FUNCTION_BLOCK GATE_CYCLE
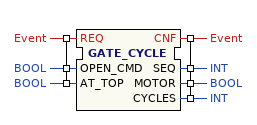
  EVENT_INPUT
    REQ WITH OPEN_CMD, AT_TOP;
  END_EVENT
  EVENT_OUTPUT
    CNF WITH SEQ, MOTOR, CYCLES;
  END_EVENT
  VAR_INPUT
    OPEN_CMD : BOOL;
    AT_TOP : BOOL;
  END_VAR
  VAR_OUTPUT
    SEQ : INT;
    MOTOR : BOOL;
    CYCLES : INT;
  END_VAR
  VAR
    SEQ_STATE : INT;
    SEQ_START_TIME : TIME;
  END_VAR
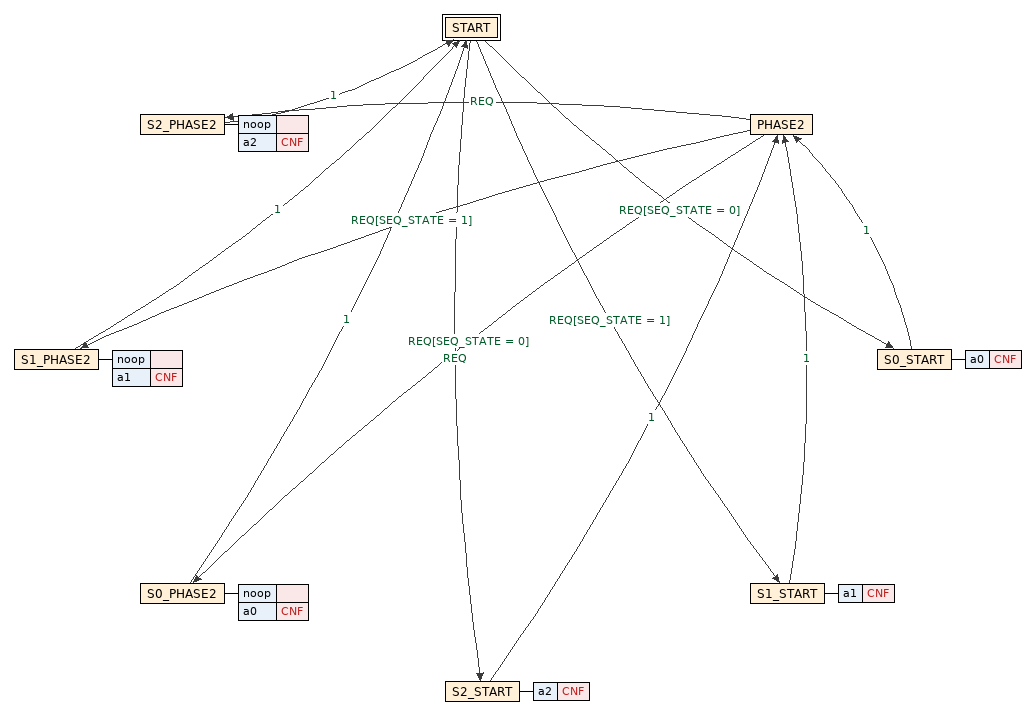
  EC_STATES
    START;
    PHASE2;
    S0_START : a0 -> CNF;
    S1_START : a1 -> CNF;
    S2_START : a2 -> CNF;
    S0_PHASE2 : noop, a0 -> CNF;
    S1_PHASE2 : noop, a1 -> CNF;
    S2_PHASE2 : noop, a2 -> CNF;
  END_STATES
  EC_TRANSITIONS
    START TO S0_START := REQ[SEQ_STATE = 0];
    START TO S1_START := REQ[SEQ_STATE = 1];
    START TO S2_START := REQ;
    PHASE2 TO S0_PHASE2 := REQ[SEQ_STATE = 0];
    PHASE2 TO S1_PHASE2 := REQ[SEQ_STATE = 1];
    PHASE2 TO S2_PHASE2 := REQ;
    S0_START TO PHASE2 := 1;
    S1_START TO PHASE2 := 1;
    S2_START TO PHASE2 := 1;
    S0_PHASE2 TO START := 1;
    S1_PHASE2 TO START := 1;
    S2_PHASE2 TO START := 1;
  END_TRANSITIONS
  ALGORITHM a0 IN ST:
MOTOR := FALSE;
IF OPEN_CMD THEN SEQ := 1; END_IF;
SEQ_STATE := SEQ;
  END_ALGORITHM
  ALGORITHM a1 IN ST:
MOTOR := TRUE;
IF AT_TOP THEN SEQ := 2; END_IF;
SEQ_STATE := SEQ;
  END_ALGORITHM
  ALGORITHM a2 IN ST:
MOTOR := FALSE;
CYCLES := CYCLES + 1;
SEQ := 0;
SEQ_STATE := SEQ;
  END_ALGORITHM
  ALGORITHM noop IN ST:
CYCLES := CYCLES;
  END_ALGORITHM
END_FUNCTION_BLOCK
